SUBAPPLICATION AR_GT_0 (* Prüft ob AR-Adapter Wert > 0.0 ist (AX-Adapter Ausgang) - analog AX_GT_0_UINT, aber fuer adapter-native AR_GT (2 AR-Sockets) statt REQ/CNF-F_GT: die feste Vergleichskonstante 0.0 kann bei einem Adapter-Socket nicht als FB-Parameter gesetzt werden, deshalb intern ueber LIT_0 (initval_AR) eingespeist. Kapselt dieses Muster, damit Aufrufer nicht jedes Mal selbst einen LIT_0-FB anlegen und verdrahten muessen (Franz: 'AR_GT_Aktiv kreuzt die beiden Eingaenge'). *)
  (* Standard: 61499-2; Description: Copyright (c) 2026 Büngener Schuder GmbH This program and the accompanying materials are made available under the terms of the Eclipse Public License 2.0 which is available at https://www.eclipse.org/legal/epl-2.0/ SPDX-License-Identifier: EPL-2.0 *)
  (* Version 1.0, 2026-10-15, Franz Höpfinger, Büngener Schuder GmbH, initial implementation - aus Aufnahme_PVEA/Igelband_PVEA/Elevator_PVEA.SUB herausgeloest (dort AR_GT_Aktiv+LIT_0 jeweils einzeln verdrahtet, mit sich kreuzenden Leitungen in der IDE-Ansicht). *)
  PACKAGE MyLib::sys;
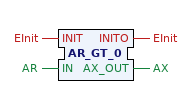
  EVENT_INPUT
    INIT : EInit; (* Initialization Request *)
  END_EVENT
  EVENT_OUTPUT
    INITO : EInit; (* Initialization Confirm *)
  END_EVENT
  SOCKETS
    IN : adapter::types::unidirectional::AR; (* Wert, der gegen 0.0 verglichen wird *)
  END_SOCKETS
  PLUGS
    AX_OUT : adapter::types::unidirectional::AX; (* TRUE wenn IN > 0.0 *)
  END_PLUGS
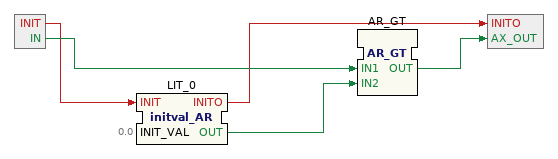
  FBS
    LIT_0 : adapter::types::unidirectional::AR::initval::initval_AR(INIT_VAL := 0.0);
    AR_GT : adapter::iec61131::comparison::AR_GT;
  END_FBS
  EVENT_CONNECTIONS
    INIT TO LIT_0.INIT;
    LIT_0.INITO TO INITO;
  END_CONNECTIONS
  ADAPTER_CONNECTIONS
    IN TO AR_GT.IN1;
    LIT_0.OUT TO AR_GT.IN2;
    AR_GT.OUT TO AX_OUT;
  END_CONNECTIONS
END_SUBAPPLICATION
